TYPE E_PortalState_New :
(
	eInit := 0,
	eIdle,
	eSetJob,
	eOpenGripper,
	eCloseGripper,
	eError,
	eMoveToStone,
	eTrspStone,
	eStampTriggered,
	eHome,
	eEStop,
	eAfterEStop,
	eManualMode,
	eDebug
);
END_TYPE

(* stored: Version 1.1.0.1, ProductVersion 3.1.4024.12
   DUT E_PortalState_New: Id {2ffab6f6-1ac0-491d-b991-c6eb365772ff} *)
